PROGRAM FunktionBlockDiagram
VAR
	ixLevel : INT;
	mxHighLevel : BOOL;
	mxLowerLevel : BOOL;
	mxLevel : INT;
	
	miProportional : INT := 10;
	miConst : INT := 50;
	miNewProp :  INT;
	
	msNormalLevel : STRING  := 'Normal Level';
	msHighLevel : STRING := 'High Level';
	msLowerLevel : STRING := 'Lower Level';
	
	
END_VAR

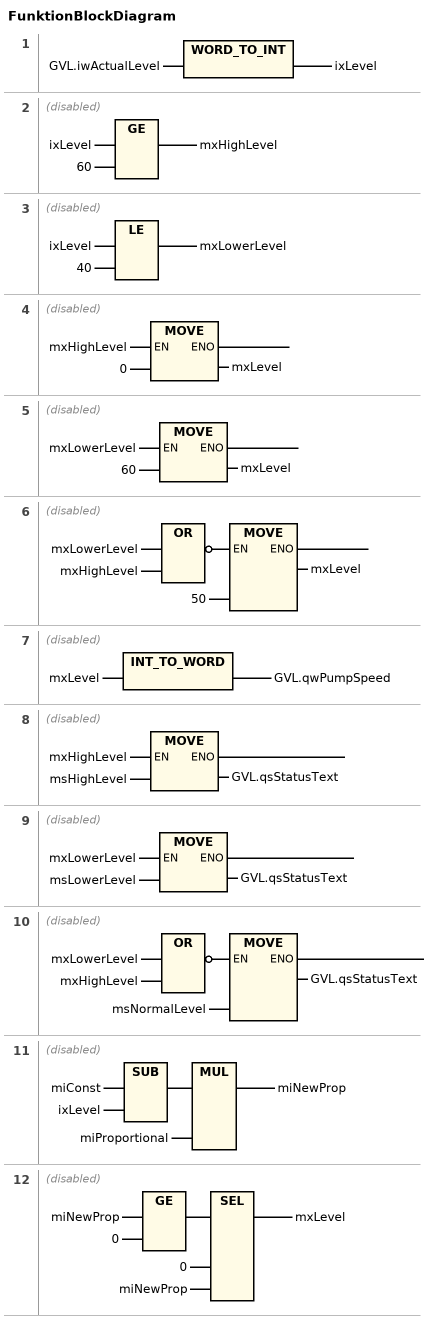
// NETWORK 1
ixLevel := WORD_TO_INT(GVL.iwActualLevel);

// NETWORK 2 (disabled)
// mxHighLevel := ixLevel >= 60;

// NETWORK 3 (disabled)
// mxLowerLevel := ixLevel <= 40;

// NETWORK 4 (disabled)
// IF mxHighLevel THEN mxLevel := 0; END_IF

// NETWORK 5 (disabled)
// IF mxLowerLevel THEN mxLevel := 60; END_IF

// NETWORK 6 (disabled)
// IF NOT (mxLowerLevel OR mxHighLevel) THEN mxLevel := 50; END_IF

// NETWORK 7 (disabled)
// GVL.qwPumpSpeed := INT_TO_WORD(mxLevel);

// NETWORK 8 (disabled)
// IF mxHighLevel THEN GVL.qsStatusText := msHighLevel; END_IF

// NETWORK 9 (disabled)
// IF mxLowerLevel THEN GVL.qsStatusText := msLowerLevel; END_IF

// NETWORK 10 (disabled)
// IF NOT (mxLowerLevel OR mxHighLevel) THEN GVL.qsStatusText := msNormalLevel; END_IF

// NETWORK 11 (disabled)
// miNewProp := (miConst - ixLevel) * miProportional;

// NETWORK 12 (disabled)
// mxLevel := SEL(miNewProp >= 0, 0, miNewProp);

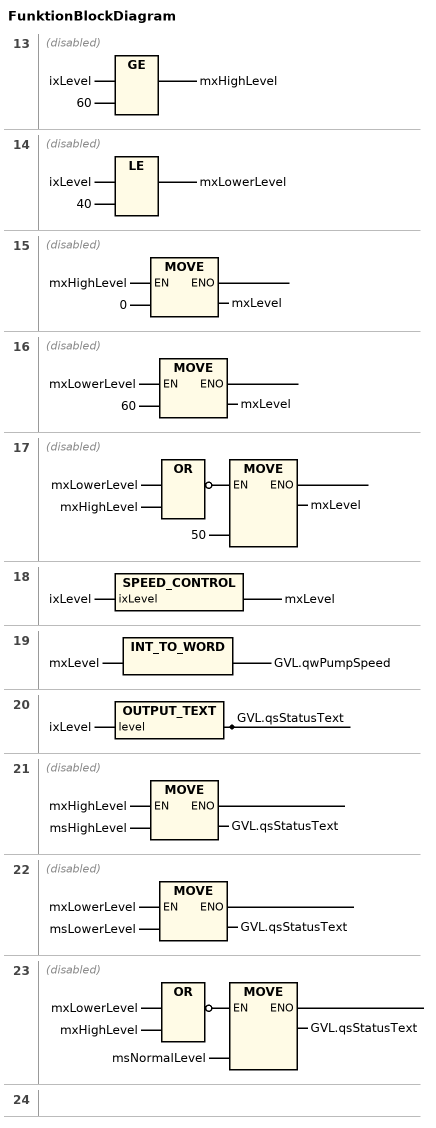
// NETWORK 13 (disabled)
// mxHighLevel := ixLevel >= 60;

// NETWORK 14 (disabled)
// mxLowerLevel := ixLevel <= 40;

// NETWORK 15 (disabled)
// IF mxHighLevel THEN mxLevel := 0; END_IF

// NETWORK 16 (disabled)
// IF mxLowerLevel THEN mxLevel := 60; END_IF

// NETWORK 17 (disabled)
// IF NOT (mxLowerLevel OR mxHighLevel) THEN mxLevel := 50; END_IF

// NETWORK 18
mxLevel := SPEED_CONTROL(ixLevel := ixLevel);

// NETWORK 19
GVL.qwPumpSpeed := INT_TO_WORD(mxLevel);

// NETWORK 20
GVL.qsStatusText := OUTPUT_TEXT(level := ixLevel);

// NETWORK 21 (disabled)
// IF mxHighLevel THEN GVL.qsStatusText := msHighLevel; END_IF

// NETWORK 22 (disabled)
// IF mxLowerLevel THEN GVL.qsStatusText := msLowerLevel; END_IF

// NETWORK 23 (disabled)
// IF NOT (mxLowerLevel OR mxHighLevel) THEN GVL.qsStatusText := msNormalLevel; END_IF

// NETWORK 24

END_PROGRAM

(* stored: Version 1.1.0.1
   POU FunktionBlockDiagram: Id {bb9f87a0-c1f0-406b-9126-1016eb4ae4b7}, SpecialFunc None *)
